{attribute 'qualified_only'}
{attribute 'strict'}
{attribute 'to_string'}
TYPE E_ULint :
(
	eOptionA := 0,
	eOptionB,
	eOptionC
) ULINT;
END_TYPE

(* stored: Version 1.1.0.1, ProductVersion 3.1.4026.19
   DUT E_ULint: Id {1816863d-06fe-47ab-9a02-1608d5227572} *)
